(*
SPDX-FileCopyrightText: © 2026 Oleksandr Tiutyk <trofimich@gmail.com>
SPDX-License-Identifier: MIT
License: https://opensource.org/license/mit
*)

(*!
<summary>Checks that an incomplete child enters INVALID after its initialization timeout.</summary>
<description>
Owns a fresh simulated automation fixture and advances one initialization call per PLC cycle.
The fixture limits attempts to fifty calls. No native resources or hardware are involved.
</description>
*)

{attribute 'no_assign'}
{attribute 'no_explicit_call' := 'do not call this function block directly'}
FUNCTION_BLOCK AutomationChildInitializationTimeoutTest EXTENDS TOF_Testing.MultiCycleTest
VAR_STAT
	{attribute 'hide'}
	_ClassName : STRING := __POUNAME();
END_VAR
VAR
	_Fixture : POINTER TO AutomationComponentTestFixture;
END_VAR

(*!
<summary>Creates the fixture, whose attempt limit bounds the scenario.</summary>
*)
METHOD PROTECTED BeforeTest
_Timeout := T#0S;
_Fixture := __NEW(AutomationComponentTestFixture);

IF _Fixture = 0 THEN
	TOF_Core.DynamicMemoryManager.RaiseAllocationFailure();
END_IF
END_METHOD

(*!
<summary>Advances one child initialization call and reports completion when the result is observable.</summary>
*)
METHOD PROTECTED ExecuteTest : TOF_Testing.TEST_CYCLE_RESULT
VAR
	assertions : REFERENCE TO TOF_Testing.Assertions;
END_VAR
assertions REF= Assert;
ExecuteTest := _Fixture^.AdvanceInitializationTimeout(assertions := assertions);
END_METHOD

(*!
<summary>Releases the fixture before publishing the result, after success or failure.</summary>
*)
METHOD PROTECTED AfterTest
VAR
	fixture : POINTER TO AutomationComponentTestFixture;
END_VAR
fixture := _Fixture;
_Fixture := 0;

IF fixture <> 0 THEN
	__DELETE(fixture);
END_IF
END_METHOD

(*!
<summary>Releases a still-owned fixture when the case is unloaded.</summary>
<param name="bInCopyCode">TwinCAT copy-code exit marker. Leave copied ownership with the new instance.</param>
*)
METHOD FB_exit : BOOL
VAR_INPUT
	bInCopyCode : BOOL;
END_VAR
IF NOT bInCopyCode AND_THEN _Fixture <> 0 THEN
	__DELETE(_Fixture);
END_IF

FB_exit := TRUE;
END_METHOD

(*!
<summary>Borrows the concrete class name. Callers must not modify it.</summary>
*)
{attribute 'monitoring' := 'call'}
PROPERTY ClassName : REFERENCE TO STRING
GET
ClassName REF= _ClassName;
END_GET
END_PROPERTY

(*!
<summary>Borrows the project namespace name. Callers must not modify it.</summary>
*)
{attribute 'monitoring' := 'call'}
PROPERTY NamespaceName : REFERENCE TO STRING
GET
NamespaceName REF= CurrentNamespace.Name;
END_GET
END_PROPERTY

(*!
<summary>Reports the complete instance size in bytes.</summary>
*)
{attribute 'monitoring' := 'call'}
PROPERTY SelfSize : ULINT
GET
SelfSize := XSIZEOF(THIS^);
END_GET
END_PROPERTY

END_FUNCTION_BLOCK

(* stored: Version 1.1.0.1
   POU AutomationChildInitializationTimeoutTest: Id {ef66d2a6-ff4f-4fc7-af7b-b467f210ddab}, SpecialFunc None
   Method BeforeTest: Id {ad56f804-69d2-4d2b-92db-e2ed7851b84d}
   Method ExecuteTest: Id {68ce8353-07ce-46f5-a2a9-eaf2157cff2a}
   Method AfterTest: Id {8bbc3447-c73b-4ecf-8cd3-a07b1b6ef66e}
   Method FB_exit: Id {e86534fa-61d7-418b-942f-01669a6f3a99}
   Property ClassName: Id {f9034aa0-fe7f-4026-892a-f0019c2aa13d}
   Get Get: Id {35b5c624-e1ec-4a4a-a1f6-25f59f519340}
   Property NamespaceName: Id {7e6c6592-ed82-4975-b9f3-bda648ba45d9}
   Get Get: Id {9ae8a4f7-95fa-46c9-a12f-d8a92ccc7931}
   Property SelfSize: Id {50199e84-22dc-4b75-b41f-a85c79acb177}
   Get Get: Id {d0fd14b8-c0e1-48aa-891b-3e2d46ddfa15} *)
